                                                   #SUBSEQUENT_ENCODING:  // Statement section case 2 to 4
                                                       FOR #tempLoopCounter := #statClientIdPos TO LEN(#clientIdentifier) DO
                                                           "LMQTT_ConvertToUtf8"(character := #clientIdentifier[#tempLoopCounter],
                                                                                 convertedUtf8 => #tempConvertedUtf8,
                                                                                 bytesUsed => #tempBytesUsedUtf8,
                                                                                 error => #tempErrorConvertUtf8,
                                                                                 status => #tempStatusConvertUtf8);
                                                           IF #statSendBufferPos + #tempBytesUsedUtf8 <= #MAX_BUFFER_LEN_SEND THEN
                                                               #statClientIdPos += 1;
                                                               CASE #tempBytesUsedUtf8 OF
                                                                   #UTF_1_BYTE_USED:  // Statement section case 1
                                                                       #statSendBuffer[#statSendBufferPos] := #tempConvertedUtf8.%B0;
                                                                       #statSendBufferPos += 1;
                                                                   #UTF_2_BYTE_USED:
                                                                       #statSendBuffer[#statSendBufferPos] := #tempConvertedUtf8.%B0;
                                                                       #statSendBufferPos += 1;
                                                                       #statSendBuffer[#statSendBufferPos] := #tempConvertedUtf8.%B1;
                                                                       #statSendBufferPos += 1;
                                                                   #UTF_3_BYTE_USED:  // Statement section case 2 to 4
                                                                       #statSendBuffer[#statSendBufferPos] := #tempConvertedUtf8.%B0;
                                                                       #statSendBufferPos += 1;
                                                                       #statSendBuffer[#statSendBufferPos] := #tempConvertedUtf8.%B1;
                                                                       #statSendBufferPos += 1;
                                                                       #statSendBuffer[#statSendBufferPos] := #tempConvertedUtf8.%B2;
                                                                       #statSendBufferPos += 1;
                                                                   ELSE  // Statement section ELSE
                                                                       ;
                                                               END_CASE;
                                                           ELSE
                                                               // When buffer full
                                                               EXIT;
                                                           END_IF;
                                                       END_FOR;
                                                       IF #statClientIdPos >= LEN(#clientIdentifier) THEN
                                                           #statClientIdEncodeState := #ENCODE_DONE;
                                                       END_IF;
                                                   ELSE  // Statement section ELSE
                                                       ; // IDLE / SKIP
                                               END_CASE;
                                           END_IF;

                                           // Will Topic
                                           // If the Will Flag is set to 1, the Will Topic is the next field in the payload. It must be > 0 Bytes

                                           IF #statClientIdEncodeState = #ENCODE_DONE
                                               AND #statSendBufferPos <= #MAX_BUFFER_LEN_SEND - #TWO_BYTE_LEN_INFO THEN
                                               // When Client Id is encoded and buffer not full
                                               // And willTopic is used
                                               CASE #statWillTopicEncodeState OF
                                                   #FIRST_ENCODING:  // Statement section case 1
                                                       // ADD len info into packet

                                                       #tempWordForSliceAddress := UINT_TO_WORD(#statWillTopicLenUtf8Encoded);
                                                       #statSendBuffer[#statSendBufferPos] := #tempWordForSliceAddress.%B1; // MSB
                                                       #statSendBufferPos += 1;
                                                       #statSendBuffer[#statSendBufferPos] := #tempWordForSliceAddress.%B0; // LSB
                                                       #statSendBufferPos += 1;

                                                       FOR #tempLoopCounter := #statWillTopicPos TO LEN(#willtopic) DO
                                                           "LMQTT_ConvertToUtf8"(character := #willtopic[#tempLoopCounter],
                                                                                 convertedUtf8 => #tempConvertedUtf8,
                                                                                 bytesUsed => #tempBytesUsedUtf8,
                                                                                 error => #tempErrorConvertUtf8,
                                                                                 status => #tempStatusConvertUtf8);

                                                           IF #statSendBufferPos + #tempBytesUsedUtf8 <= #MAX_BUFFER_LEN_SEND THEN
                                                               // Increment when successful
                                                               #statWillTopicPos += 1;

                                                               CASE #tempBytesUsedUtf8 OF
                                                                   #UTF_1_BYTE_USED:  // Statement section case 1
                                                                       #statSendBuffer[#statSendBufferPos] := #tempConvertedUtf8.%B0;
                                                                       #statSendBufferPos += 1;
                                                                   #UTF_2_BYTE_USED:
                                                                       #statSendBuffer[#statSendBufferPos] := #tempConvertedUtf8.%B0;
                                                                       #statSendBufferPos += 1;
                                                                       #statSendBuffer[#statSendBufferPos] := #tempConvertedUtf8.%B1;
                                                                       #statSendBufferPos += 1;
                                                                   #UTF_3_BYTE_USED:  // Statement section case 2 to 4
                                                                       #statSendBuffer[#statSendBufferPos] := #tempConvertedUtf8.%B0;
                                                                       #statSendBufferPos += 1;
                                                                       #statSendBuffer[#statSendBufferPos] := #tempConvertedUtf8.%B1;
                                                                       #statSendBufferPos += 1;
                                                                       #statSendBuffer[#statSendBufferPos] := #tempConvertedUtf8.%B2;
                                                                       #statSendBufferPos += 1;
                                                                   ELSE  // Statement section ELSE
                                                                       ;
                                                               END_CASE;
                                                           ELSE
                                                               // When buffer full
                                                               #statWillTopicEncodeState := #SUBSEQUENT_ENCODING;
                                                               EXIT;
                                                           END_IF;
                                                       END_FOR;

                                                       IF #statWillTopicPos >= LEN(#willtopic) THEN
                                                           #statWillTopicEncodeState := #ENCODE_DONE;
                                                       END_IF;

                                                   #SUBSEQUENT_ENCODING:  // Statement section case 2 to 4
                                                       FOR #tempLoopCounter := #statWillTopicPos TO LEN(#willtopic) DO
                                                           "LMQTT_ConvertToUtf8"(character := #willtopic[#tempLoopCounter],
                                                                                 convertedUtf8 => #tempConvertedUtf8,
                                                                                 bytesUsed => #tempBytesUsedUtf8,
                                                                                 error => #tempErrorConvertUtf8,
                                                                                 status => #tempStatusConvertUtf8);

                                                           IF #statSendBufferPos + #tempBytesUsedUtf8 <= #MAX_BUFFER_LEN_SEND THEN
                                                               #statWillTopicPos += 1;
                                                               CASE #tempBytesUsedUtf8 OF
                                                                   #UTF_1_BYTE_USED:  // Statement section case 1
                                                                       #statSendBuffer[#statSendBufferPos] := #tempConvertedUtf8.%B0;
                                                                       #statSendBufferPos += 1;
                                                                   #UTF_2_BYTE_USED:
                                                                       #statSendBuffer[#statSendBufferPos] := #tempConvertedUtf8.%B0;
                                                                       #statSendBufferPos += 1;
                                                                       #statSendBuffer[#statSendBufferPos] := #tempConvertedUtf8.%B1;
                                                                       #statSendBufferPos += 1;
                                                                   #UTF_3_BYTE_USED:  // Statement section case 2 to 4
                                                                       #statSendBuffer[#statSendBufferPos] := #tempConvertedUtf8.%B0;
                                                                       #statSendBufferPos += 1;
                                                                       #statSendBuffer[#statSendBufferPos] := #tempConvertedUtf8.%B1;
                                                                       #statSendBufferPos += 1;
                                                                       #statSendBuffer[#statSendBufferPos] := #tempConvertedUtf8.%B2;
                                                                       #statSendBufferPos += 1;
                                                                   ELSE  // Statement section ELSE
                                                                       ;
                                                               END_CASE;
                                                           ELSE
                                                               // When buffer full
                                                               EXIT;
                                                           END_IF;
                                                       END_FOR;
                                                       IF #statWillTopicPos >= LEN(#willtopic) THEN
                                                           #statWillTopicEncodeState := #ENCODE_DONE;
                                                       END_IF;

                                                   ELSE  // Statement section ELSE
                                                       ;
                                               END_CASE;
                                           END_IF;

                                           // Will Message
                                           // This field consists OF a two Byte length followed BY the payload FOR the Will message expressed as a sequence bytes.

                                           IF #statClientIdEncodeState = #ENCODE_DONE
                                               AND #statWillTopicEncodeState = #ENCODE_DONE
                                               AND #statSendBufferPos <= #MAX_BUFFER_LEN_SEND - #TWO_BYTE_LEN_INFO THEN
                                               // When Client Id is encoded and buffer not full
                                               CASE #statWillMessageEncodeState OF
                                                   #FIRST_ENCODING:  // Statement section case 1
                                                       // ADD len info into packet

                                                       #tempWordForSliceAddress := UINT_TO_WORD(#statWillMessageCnt);
                                                       #statSendBuffer[#statSendBufferPos] := #tempWordForSliceAddress.%B1; // MSB
                                                       #statSendBufferPos += 1;
                                                       #statSendBuffer[#statSendBufferPos] := #tempWordForSliceAddress.%B0; // LSB
                                                       #statSendBufferPos += 1;

                                                       #tempLowerWillMsgArrayBoundary := LOWER_BOUND(ARR := #willMsgPayload, DIM := #ONE_DIMENSION);

                                                       IF #statWillMessageCnt > 0 THEN // will message exists
                                                           FOR #tempLoopCounter := #statWillMessagePos TO UINT_TO_DINT(#statWillMessageCnt - 1) DO
                                                               IF #statSendBufferPos <= #MAX_BUFFER_LEN_SEND THEN
                                                                   #statSendBuffer[#statSendBufferPos] := #willMsgPayload[#tempLowerWillMsgArrayBoundary + #tempLoopCounter];
                                                                   #statSendBufferPos += 1;
                                                                   // Increment when successful
                                                                   #statWillMessagePos += 1;
                                                               ELSE
                                                                   // When buffer full
                                                                   #statWillMessageEncodeState := #SUBSEQUENT_ENCODING;
                                                                   EXIT;
                                                               END_IF;
                                                           END_FOR;
                                                       END_IF;

                                                       // If everything was copied successfull
                                                       IF #statWillMessagePos >= #statWillMessageCnt THEN
                                                           #statWillMessageEncodeState := #ENCODE_DONE;
                                                       END_IF;

                                                   #SUBSEQUENT_ENCODING:  // Statement section case 2 to 4
                                                       #tempLowerWillMsgArrayBoundary := LOWER_BOUND(ARR := #willMsgPayload, DIM := #ONE_DIMENSION);

                                                       FOR #tempLoopCounter := #statWillMessagePos TO UINT_TO_DINT(#statWillMessageCnt - 1) DO
                                                           IF #statSendBufferPos <= #MAX_BUFFER_LEN_SEND THEN
                                                               #statSendBuffer[#statSendBufferPos] := #willMsgPayload[#tempLowerWillMsgArrayBoundary + #tempLoopCounter];
                                                               #statSendBufferPos += 1;
                                                               // Increment when successful
                                                               #statWillMessagePos += 1;
                                                           ELSE
                                                               // When Buffer Full
                                                               EXIT;
                                                           END_IF;
                                                       END_FOR;
                                                       // If everything was copied successfull
                                                       IF #statWillMessagePos >= #statWillMessageCnt THEN
                                                           #statWillMessageEncodeState := #ENCODE_DONE;
                                                       END_IF;


                                                   ELSE  // Statement section ELSE
                                                       ;
                                               END_CASE;
                                           END_IF;

                                           // Username
                                           // If the Username Flag is set to 1, the Username the next field in the payload. It must be > 0 Bytes

                                           IF #statClientIdEncodeState = #ENCODE_DONE
                                               AND (#statWillTopicEncodeState = #ENCODE_DONE OR #statWillTopicEncodeState = #NOT_USED_NO_ENCODING)
                                               AND (#statWillMessageEncodeState = #ENCODE_DONE OR #statWillTopicEncodeState = #NOT_USED_NO_ENCODING)
                                               AND #statSendBufferPos <= #MAX_BUFFER_LEN_SEND - #TWO_BYTE_LEN_INFO THEN
                                               // When Will Topic and Will Message is encoded and buffer not full
                                               CASE #statUserNameEncodeState OF
                                                   #FIRST_ENCODING:  // Statement section case 1
                                                       // ADD len info into packet

                                                       #tempWordForSliceAddress := UINT_TO_WORD(#statUsernameLenUtf8Encoded);
                                                       #statSendBuffer[#statSendBufferPos] := #tempWordForSliceAddress.%B1; // MSB
                                                       #statSendBufferPos += 1;
                                                       #statSendBuffer[#statSendBufferPos] := #tempWordForSliceAddress.%B0; // LSB
                                                       #statSendBufferPos += 1;

                                                       FOR #tempLoopCounter := #statUserNamePos TO LEN(#username) DO
                                                           "LMQTT_ConvertToUtf8"(character := #username[#tempLoopCounter],
                                                                                 convertedUtf8 => #tempConvertedUtf8,
                                                                                 bytesUsed => #tempBytesUsedUtf8,
                                                                                 error => #tempErrorConvertUtf8,
                                                                                 status => #tempStatusConvertUtf8);

                                                           IF #statSendBufferPos + #tempBytesUsedUtf8 <= #MAX_BUFFER_LEN_SEND THEN
                                                               // Increment when successful
                                                               #statUserNamePos += 1;

                                                               CASE #tempBytesUsedUtf8 OF
                                                                   #UTF_1_BYTE_USED:  // Statement section case 1
                                                                       #statSendBuffer[#statSendBufferPos] := #tempConvertedUtf8.%B0;
                                                                       #statSendBufferPos += 1;
                                                                   #UTF_2_BYTE_USED:
                                                                       #statSendBuffer[#statSendBufferPos] := #tempConvertedUtf8.%B0;
                                                                       #statSendBufferPos += 1;
                                                                       #statSendBuffer[#statSendBufferPos] := #tempConvertedUtf8.%B1;
                                                                       #statSendBufferPos += 1;
                                                                   #UTF_3_BYTE_USED:  // Statement section case 2 to 4
                                                                       #statSendBuffer[#statSendBufferPos] := #tempConvertedUtf8.%B0;
                                                                       #statSendBufferPos += 1;
                                                                       #statSendBuffer[#statSendBufferPos] := #tempConvertedUtf8.%B1;
                                                                       #statSendBufferPos += 1;
                                                                       #statSendBuffer[#statSendBufferPos] := #tempConvertedUtf8.%B2;
                                                                       #statSendBufferPos += 1;
                                                                   ELSE  // Statement section ELSE
                                                                       ;
                                                               END_CASE;
                                                           ELSE
                                                               // When buffer full
                                                               #statUserNameEncodeState := #SUBSEQUENT_ENCODING;
                                                               EXIT;
                                                           END_IF;
                                                       END_FOR;

                                                       IF #statUserNamePos >= LEN(#username) THEN
                                                           #statUserNameEncodeState := #ENCODE_DONE;
                                                       END_IF;

                                                   #SUBSEQUENT_ENCODING:  // Statement section case 2 to 4
                                                       FOR #tempLoopCounter := #statUserNamePos TO LEN(#username) DO
                                                           "LMQTT_ConvertToUtf8"(character := #username[#tempLoopCounter],
                                                                                 convertedUtf8 => #tempConvertedUtf8,
                                                                                 bytesUsed => #tempBytesUsedUtf8,
                                                                                 error => #tempErrorConvertUtf8,
                                                                                 status => #tempStatusConvertUtf8);

                                                           IF #statSendBufferPos + #tempBytesUsedUtf8 <= #MAX_BUFFER_LEN_SEND THEN
                                                               #statUserNamePos += 1;
                                                               CASE #tempBytesUsedUtf8 OF
                                                                   #UTF_1_BYTE_USED:  // Statement section case 1
                                                                       #statSendBuffer[#statSendBufferPos] := #tempConvertedUtf8.%B0;
                                                                       #statSendBufferPos += 1;
                                                                   #UTF_2_BYTE_USED:
                                                                       #statSendBuffer[#statSendBufferPos] := #tempConvertedUtf8.%B0;
                                                                       #statSendBufferPos += 1;
                                                                       #statSendBuffer[#statSendBufferPos] := #tempConvertedUtf8.%B1;
                                                                       #statSendBufferPos += 1;
                                                                   #UTF_3_BYTE_USED:  // Statement section case 2 to 4
                                                                       #statSendBuffer[#statSendBufferPos] := #tempConvertedUtf8.%B0;
                                                                       #statSendBufferPos += 1;
                                                                       #statSendBuffer[#statSendBufferPos] := #tempConvertedUtf8.%B1;
                                                                       #statSendBufferPos += 1;
                                                                       #statSendBuffer[#statSendBufferPos] := #tempConvertedUtf8.%B2;
                                                                       #statSendBufferPos += 1;
                                                                   ELSE  // Statement section ELSE
                                                                       ;
                                                               END_CASE;
                                                           ELSE
                                                               // When buffer full
                                                               EXIT;
                                                           END_IF;
                                                       END_FOR;
                                                       IF #statUserNamePos >= LEN(#username) THEN
                                                           #statUserNameEncodeState := #ENCODE_DONE;
                                                       END_IF;

                                                   ELSE  // Statement section ELSE
                                                       ;
                                               END_CASE;
                                           END_IF;

                                           // Password
                                           // If the Password Flag is set to 1, the Password the next field in the payload. It must be > 0 Bytes
                                           // Password field contains 0 to 65535 bytes OF binary data prefixed with a two Byte length field which indicates the number OF bytes used

                                           IF #statClientIdEncodeState = #ENCODE_DONE
                                               AND (#statWillTopicEncodeState = #ENCODE_DONE OR #statWillTopicEncodeState = #NOT_USED_NO_ENCODING)
                                               AND (#statWillMessageEncodeState = #ENCODE_DONE OR #statWillMessageEncodeState = #NOT_USED_NO_ENCODING)
                                               AND (#statUserNameEncodeState = #ENCODE_DONE OR #statUserNameEncodeState = #NOT_USED_NO_ENCODING)
                                               AND #statSendBufferPos <= #MAX_BUFFER_LEN_SEND - #TWO_BYTE_LEN_INFO THEN
                                               // When Will Topic and Will Message is encoded and buffer not full
                                               CASE #statPasswordEncodeState OF
                                                   #FIRST_ENCODING:  // Statement section case 1
                                                       // ADD len info into packet

                                                       #tempWordForSliceAddress := UINT_TO_WORD(#statPasswordLenUtf8Encoded);
                                                       #statSendBuffer[#statSendBufferPos] := #tempWordForSliceAddress.%B1; // MSB
                                                       #statSendBufferPos += 1;
                                                       #statSendBuffer[#statSendBufferPos] := #tempWordForSliceAddress.%B0; // LSB
                                                       #statSendBufferPos += 1;

                                                       FOR #tempLoopCounter := #statPasswordPos TO LEN(#password) DO
                                                           "LMQTT_ConvertToUtf8"(character := #password[#tempLoopCounter],
                                                                                 convertedUtf8 => #tempConvertedUtf8,
                                                                                 bytesUsed => #tempBytesUsedUtf8,
                                                                                 error => #tempErrorConvertUtf8,
                                                                                 status => #tempStatusConvertUtf8);

                                                           IF #statSendBufferPos + #tempBytesUsedUtf8 <= #MAX_BUFFER_LEN_SEND THEN
                                                               // Increment when successful
                                                               #statPasswordPos += 1;

                                                               CASE #tempBytesUsedUtf8 OF
                                                                   #UTF_1_BYTE_USED:  // Statement section case 1
                                                                       #statSendBuffer[#statSendBufferPos] := #tempConvertedUtf8.%B0;
                                                                       #statSendBufferPos += 1;
                                                                   #UTF_2_BYTE_USED:
                                                                       #statSendBuffer[#statSendBufferPos] := #tempConvertedUtf8.%B0;
                                                                       #statSendBufferPos += 1;
                                                                       #statSendBuffer[#statSendBufferPos] := #tempConvertedUtf8.%B1;
                                                                       #statSendBufferPos += 1;
                                                                   #UTF_3_BYTE_USED:  // Statement section case 2 to 4
                                                                       #statSendBuffer[#statSendBufferPos] := #tempConvertedUtf8.%B0;
                                                                       #statSendBufferPos += 1;
                                                                       #statSendBuffer[#statSendBufferPos] := #tempConvertedUtf8.%B1;
                                                                       #statSendBufferPos += 1;
                                                                       #statSendBuffer[#statSendBufferPos] := #tempConvertedUtf8.%B2;
                                                                       #statSendBufferPos += 1;
                                                                   ELSE  // Statement section ELSE
                                                                       ;
                                                               END_CASE;
                                                           ELSE
                                                               // When buffer full
                                                               #statPasswordEncodeState := #SUBSEQUENT_ENCODING;
                                                               EXIT;
                                                           END_IF;
                                                       END_FOR;

                                                       IF #statPasswordPos >= LEN(#password) THEN
                                                           #statPasswordEncodeState := #ENCODE_DONE;
                                                       END_IF;

                                                   #SUBSEQUENT_ENCODING:  // Statement section case 2 to 4
                                                       FOR #tempLoopCounter := #statPasswordPos TO LEN(#password) DO
                                                           "LMQTT_ConvertToUtf8"(character := #password[#tempLoopCounter],
                                                                                 convertedUtf8 => #tempConvertedUtf8,
                                                                                 bytesUsed => #tempBytesUsedUtf8,
                                                                                 error => #tempErrorConvertUtf8,
                                                                                 status => #tempStatusConvertUtf8);

                                                           IF #statSendBufferPos + #tempBytesUsedUtf8 <= #MAX_BUFFER_LEN_SEND THEN
                                                               #statPasswordPos += 1;
                                                               CASE #tempBytesUsedUtf8 OF
                                                                   #UTF_1_BYTE_USED:  // Statement section case 1
                                                                       #statSendBuffer[#statSendBufferPos] := #tempConvertedUtf8.%B0;
                                                                       #statSendBufferPos += 1;
                                                                   #UTF_2_BYTE_USED:
                                                                       #statSendBuffer[#statSendBufferPos] := #tempConvertedUtf8.%B0;
                                                                       #statSendBufferPos += 1;
                                                                       #statSendBuffer[#statSendBufferPos] := #tempConvertedUtf8.%B1;
                                                                       #statSendBufferPos += 1;
                                                                   #UTF_3_BYTE_USED:  // Statement section case 2 to 4
                                                                       #statSendBuffer[#statSendBufferPos] := #tempConvertedUtf8.%B0;
                                                                       #statSendBufferPos += 1;
                                                                       #statSendBuffer[#statSendBufferPos] := #tempConvertedUtf8.%B1;
                                                                       #statSendBufferPos += 1;
                                                                       #statSendBuffer[#statSendBufferPos] := #tempConvertedUtf8.%B2;
                                                                       #statSendBufferPos += 1;
                                                                   ELSE  // Statement section ELSE
                                                                       ;
                                                               END_CASE;
                                                           ELSE
                                                               // When buffer full
                                                               EXIT;
                                                           END_IF;
                                                       END_FOR;
                                                       IF #statPasswordPos >= LEN(#password) THEN
                                                           #statPasswordEncodeState := #ENCODE_DONE;
                                                       END_IF;

                                                   ELSE  // Statement section ELSE
                                                       ;
                                               END_CASE;
                                           END_IF;

                                           // set Sendlen for TSendC Block
                                           #statTsendcLen := #statSendBufferPos; // Buffer pos equals amount of elements in send array
                                           // reset buffer pos
                                           #statSendBufferPos := 0;
                                           // enable Send Req
                                           #statTsendcReq := TRUE;
                                           // Set Watchdog
                                           #statEnableTimerCommandWatchdog := TRUE;
                                           // wait for send to be done
                                           #statMqttConnectState := #MQTT_CONNECT_STATE_SEND_PACKET_WAIT_FOR_CONNACK;
                                       END_IF;
                                   END_REGION BUILD_CONNECT_PACKET

                               #MQTT_CONNECT_STATE_SEND_PACKET_WAIT_FOR_CONNACK:
                                   REGION SEND_CONNECT_PACKET_WAIT_FOR_CONNACK
                                       // check tsend status
                                       IF NOT #tempTsendcBusy AND #tempTsendcStatus = #TSENDC_JOB_DONE THEN
                                           IF (#statClientIdEncodeState = #ENCODE_DONE OR #statClientIdEncodeState = #NOT_USED_NO_ENCODING)
                                               AND (#statWillTopicEncodeState = #ENCODE_DONE OR #statWillTopicEncodeState = #NOT_USED_NO_ENCODING)
                                               AND (#statWillMessageEncodeState = #ENCODE_DONE OR #statWillMessageEncodeState = #NOT_USED_NO_ENCODING)
                                               AND (#statUserNameEncodeState = #ENCODE_DONE OR #statUserNameEncodeState = #NOT_USED_NO_ENCODING)
                                               AND (#statPasswordEncodeState = #ENCODE_DONE OR #statPasswordEncodeState = #NOT_USED_NO_ENCODING) THEN
                                               // Encoding done all sent
                                               #statPacketHeaderEncodeDone := FALSE;
                                           ELSE
                                               // More to Encode and send
                                               #statEnableTimerCommandWatchdog := FALSE;
                                               #statMqttConnectState := #MQTT_CONNECT_STATE_BUILD_PACKET;
                                           END_IF;
                                       END_IF;

                                       // Check Connect ACK packet
                                       CASE #tempMqttConnAckRcvStatus OF
                                           #NO_RESPONSE:  // IDLE
                                               // Check watchdog
                                               IF #instTimerCommandWatchdog.Q THEN
                                                   #statEnableTimerCommandWatchdog := FALSE;
                                                   #statPacketHeaderEncodeDone := FALSE;
                                                   #statStatus := #ERR_MQTT_CONNECT_TIMEOUT; // Set correct status that identifies error clearly
                                                   #statSubfunctionStatus := #ERR_MQTT_CONNECT_TIMEOUT; // Status or return value of called FBs, FCs and system blocks
                                                   #statFBErrorState := #statFBState; // Set error state number for diagnostic 
                                                   #statErrorAutoCleared := TRUE;
                                                   #statMqttConnectState := #MQTT_CONNECT_STATE_BUILD_PACKET;
                                               END_IF;
                                           #RESPONSE_GOOD:
                                               // disable watchdog
                                               #statEnableTimerCommandWatchdog := FALSE;
                                               // Encoding done all sent
                                               #statPacketHeaderEncodeDone := FALSE;
                                               // Go to Connected
                                               #statMqttConnectState := #MQTT_CONNECT_STATE_CONNECTED;
                                               #statStatus := #STATUS_MQTT_CONNECTED;
                                       END_CASE;
                                   END_REGION REGION SEND_CONNECT_PACKET

                               #MQTT_CONNECT_STATE_CONNECTED:
                                   REGION CONNECTED
                                       // Check Rising edge of input commands
                                       #tempCommandInput.%X0 := #tempPublish AND NOT #statPublishOld;
                                       #tempCommandInput.%X1 := #tempSubscribe AND NOT #statSubscribeOld;
                                       #tempCommandInput.%X2 := #tempUnsubscribe AND NOT #statUnsubscribeOld;

                                       // Start the keepalive timer if used
                                       #statEnableMqttKeepAliveTimer := #statMqttKeepAliveUsed;

                                       // set status to connected after successfully executed job
                                       IF #statStatus = #STATUS_JOB_EXECUTED THEN
                                           #statStatus := #STATUS_MQTT_CONNECTED;
                                       END_IF;

                                       // Reset done bit
                                       IF #statDone = TRUE
                                           AND #tempPublish = FALSE
                                           AND #tempSubscribe = FALSE
                                           AND #tempUnsubscribe = FALSE
                                       THEN
                                           #statDone := FALSE;
                                       END_IF;

                                       REGION MQTT_COMMANDS
                                           // When state machine is ready for a new input then assign correct command
                                           // Ping job can be overwritten by a command.
                                           IF #tempCommandInput <> #NO_COMMAND
                                               AND (#statMqttCommandState = #MQTT_COMMAND_STATE_NO_PROCESSING OR #statMqttCommandState = #MQTT_COMMAND_STATE_SEND_PING)
                                           THEN
                                               // New Input set, reset done flag
                                               #statDone := FALSE;
                                               #statMqttCommandState := BYTE_TO_DINT(#tempCommandInput);
                                           END_IF;

                                           CASE #statMqttCommandState OF
                                               #MQTT_COMMAND_STATE_NO_PROCESSING:
                                                   // EMPTY STATE
                                                   ;
                                               #MQTT_COMMAND_STATE_BUILD_PUBLISH:  // Statement section case 1
                                                   REGION PUBLISH_TO_TOPIC
                                                       // Remaining Length is the length of the variable header (TOPIC NAME + PacketID) plus the length of the Payload. 
                                                       // Max Len of Mqtt packets is per Standard 268,435,455 Bytes (ff,ff,ff,7f)
                                                       // Calculate Remain Len will be
                                                       // Len of TOPIC   (max 3*16382 WChars= 49.146 Bytes)
                                                       // plus Len of PacketID (2 Bytes)
                                                       // plus Len of Payload (max 268,435,455 - 49.146 - 2 = 268.386.307 Bytes ca. 268 MB)
                                                       // Max Array / DB Len in TIA portal is around 16 MB or 16.777.216 Byte
                                                       // Set Status
                                                       #statStatus := #STATUS_MQTT_PUBLISH;

                                                       // Must obey, if not currently sending PubAck Msg on a subscription
                                                       // Else, try in the next cycle
                                                       IF #tempTsendcBusy = FALSE // when tsendC is ready
                                                           AND #tempTsendcDone = FALSE // tsendC did not finish in this cycle
                                                           AND #statTsendcReq = FALSE // TsendC request was not already requested by pub ack msg
                                                       THEN
                                                           IF #statPacketHeaderEncodeDone = FALSE THEN

                                                               // Init
                                                               #statSendPacketTotalRemLen := 0;
                                                               #statSendBufferPos := 0;
                                                               #statPublishQos := #qos;
                                                               #statPublishMessageCnt := #publishMsgLen;
                                                               #statPublishTopicEncodeState := #FIRST_ENCODING;
                                                               #statPublishTopicPos := #FIRST_CHARACTER;
                                                               #statPublishTopicLenUtf8Encoded := 0;
                                                               #statPacketId += 1;// increment
                                                               IF (#statPacketId = 0) THEN
                                                                   #statPacketId := 1;
                                                               END_IF;
                                                               #statPacketIdEncoded := FALSE;
                                                               #statPublishEncodeMessageState := #SUBSEQUENT_ENCODING; // No len info necessary so start directly at subsequent.
                                                               #statPublishMessagePos := 0; // first array element

                                                               // verify PayloadLen
                                                               #tempMaxPublishDataArrayLen := ABS(UPPER_BOUND(ARR := #publishMsgPayload, DIM := #ONE_DIMENSION) - LOWER_BOUND(ARR := #publishMsgPayload, DIM := #ONE_DIMENSION)) + #ARRAY_LEN_OFFSET_PLUS_1;

                                                               // check necessary boundaries
                                                               IF #tempMaxPublishDataArrayLen < #statPublishMessageCnt THEN
                                                                   #statStatus := #ERR_CNT_EXCEEDS_ARRAY_DIMENSION; // Set correct status that identifies error clearly
                                                                   #statSubfunctionStatus := #ERR_CNT_EXCEEDS_ARRAY_DIMENSION; // Status or return value of called FBs, FCs and system blocks
                                                                   #statFBErrorState := #statFBState; // Set error state number for diagnostic 
                                                                   #statErrorAutoCleared := TRUE;
                                                                   #statMqttCommandState := #MQTT_COMMAND_STATE_NO_PROCESSING;
                                                               ELSIF LEN(#mqttTopic) = #LEN_NULL THEN
                                                                   #statStatus := #ERR_MQTT_COMMAND_PUBLISH_TOPIC_INVALID; // Set correct status that identifies error clearly
                                                                   #statSubfunctionStatus := #ERR_MQTT_COMMAND_PUBLISH_TOPIC_INVALID; // Status or return value of called FBs, FCs and system blocks
                                                                   #statFBErrorState := #statFBState; // Set error state number for diagnostic 
                                                                   #statErrorAutoCleared := TRUE;
                                                                   #statMqttCommandState := #MQTT_COMMAND_STATE_NO_PROCESSING;
                                                               ELSIF #statPublishQos > #MQTT_QOS_2 THEN
                                                                   #statStatus := #ERR_QOS_INVALID; // Set correct status that identifies error clearly
                                                                   #statSubfunctionStatus := #ERR_QOS_INVALID; // Status or return value of called FBs, FCs and system blocks
                                                                   #statFBErrorState := #statFBState; // Set error state number for diagnostic 
                                                                   #statErrorAutoCleared := TRUE;
                                                                   #statMqttCommandState := #MQTT_COMMAND_STATE_NO_PROCESSING;
                                                               ELSE // All ok
                                                                   // Add amount of bytes for publish message
                                                                   #statSendPacketTotalRemLen := #statSendPacketTotalRemLen + #statPublishMessageCnt;
                                                                   // add publish  topic len
                                                                   FOR #tempLoopCounter := #FIRST_CHARACTER TO LEN(#mqttTopic) DO
                                                                       "LMQTT_ConvertToUtf8"(character := #mqttTopic[#tempLoopCounter],
                                                                                             convertedUtf8 => #tempConvertedUtf8,
                                                                                             bytesUsed => #tempBytesUsedUtf8,
                                                                                             error => #tempErrorConvertUtf8,
                                                                                             status => #tempStatusConvertUtf8);
                                                                       #statPublishTopicLenUtf8Encoded := #statPublishTopicLenUtf8Encoded + #tempBytesUsedUtf8;
                                                                   END_FOR;
                                                                   #statSendPacketTotalRemLen := #statSendPacketTotalRemLen + #statPublishTopicLenUtf8Encoded + #TWO_BYTE_LEN_INFO;

                                                                   // Build Publish Telegram
                                                                   // Fixed Header - Write Packet Type
                                                                   #statSendBuffer[#statSendBufferPos] := #MQTT_MSG_TYPE_PUBLISH;
                                                                   // Set DUP flag always to FALSE
                                                                   #statSendBuffer[#statSendBufferPos].%X3 := FALSE;
                                                                   // Set QoS Level
                                                                   CASE #statPublishQos OF
                                                                       #MQTT_QOS_0:  // Statement section case 0
                                                                           #statSendBuffer[#statSendBufferPos] := #statSendBuffer[#statSendBufferPos] OR #MQTT_MSG_QOS0;
                                                                       #MQTT_QOS_1:  // Statement section case 1
                                                                           #statSendBuffer[#statSendBufferPos] := #statSendBuffer[#statSendBufferPos] OR #MQTT_MSG_QOS1;
                                                                           // Add two byte len info for Mandatory packet ID
                                                                           #statSendPacketTotalRemLen := #statSendPacketTotalRemLen + #TWO_BYTE_LEN_INFO;
                                                                       #MQTT_QOS_2: // Statement section case 2
                                                                           #statSendBuffer[#statSendBufferPos] := #statSendBuffer[#statSendBufferPos] OR #MQTT_MSG_QOS2;
                                                                           // Add two byte len info for Mandatory packet ID
                                                                           #statSendPacketTotalRemLen := #statSendPacketTotalRemLen + #TWO_BYTE_LEN_INFO;
                                                                       ELSE
                                                                           ;
                                                                   END_CASE;
                                                                   // Set retain bit
                                                                   #statSendBuffer[#statSendBufferPos].%X0 := #retain;

                                                                   #statSendBufferPos += 1; // increment

                                                                   // Write Remaining Packet Len info 
                                                                   WHILE (#statSendPacketTotalRemLen > #DEFAULT_VALUE_ZERO)
                                                                   DO// See MQTT Spec for explanation of this calculation
                                                                       #statEncodedRemPacketLenAsByte := UDINT_TO_BYTE(#statSendPacketTotalRemLen MOD #SEND_LEN_MULTIPLIER_UDINT_128);
                                                                       #statSendPacketTotalRemLen := #statSendPacketTotalRemLen / #SEND_LEN_MULTIPLIER_UDINT_128;
                                                                       // if there are more data to encode, set the top bit of this byte
                                                                       IF #statSendPacketTotalRemLen > #DEFAULT_VALUE_ZERO THEN
                                                                           // Do this and continue while loop
                                                                           #statEncodedRemPacketLenAsByte := #statEncodedRemPacketLenAsByte OR UDINT_TO_BYTE(#SEND_LEN_MULTIPLIER_UDINT_128);
                                                                           #statSendBuffer[#statSendBufferPos] := #statEncodedRemPacketLenAsByte;
                                                                           #statSendBufferPos += 1;
                                                                       ELSE
                                                                           // do this and leave while loop
                                                                           #statSendBuffer[#statSendBufferPos] := #statEncodedRemPacketLenAsByte;
                                                                           #statSendBufferPos += 1;
                                                                       END_IF;
                                                                   END_WHILE;
                                                                   // When all done, set encode to true
                                                                   #statPacketHeaderEncodeDone := TRUE;
                                                               END_IF;
                                                           END_IF;

                                                           // Header Encoded - now Topic, PacketId and Message need to be encoded.
                                                           IF #statPacketHeaderEncodeDone = TRUE THEN

                                                               // Publish Topic
                                                               IF #statSendBufferPos <= #MAX_BUFFER_LEN_SEND - #TWO_BYTE_LEN_INFO THEN
                                                                   CASE #statPublishTopicEncodeState OF
                                                                       #FIRST_ENCODING:  // Statement section case 1
                                                                           // ADD len info into packet

                                                                           #tempWordForSliceAddress := UINT_TO_WORD(#statPublishTopicLenUtf8Encoded);
                                                                           #statSendBuffer[#statSendBufferPos] := #tempWordForSliceAddress.%B1; // MSB
                                                                           #statSendBufferPos += 1;
                                                                           #statSendBuffer[#statSendBufferPos] := #tempWordForSliceAddress.%B0; // LSB
                                                                           #statSendBufferPos += 1;

                                                                           FOR #tempLoopCounter := #statPublishTopicPos TO LEN(#mqttTopic) DO
                                                                               "LMQTT_ConvertToUtf8"(character := #mqttTopic[#tempLoopCounter],
                                                                                                     convertedUtf8 => #tempConvertedUtf8,
                                                                                                     bytesUsed => #tempBytesUsedUtf8,
                                                                                                     error => #tempErrorConvertUtf8,
                                                                                                     status => #tempStatusConvertUtf8);

                                                                               IF #statSendBufferPos + #tempBytesUsedUtf8 <= #MAX_BUFFER_LEN_SEND THEN
                                                                                   #statPublishTopicPos += 1;
                                                                                   CASE #tempBytesUsedUtf8 OF
                                                                                       #UTF_1_BYTE_USED:  // Statement section case 1
                                                                                           #statSendBuffer[#statSendBufferPos] := #tempConvertedUtf8.%B0;
                                                                                           #statSendBufferPos += 1;
                                                                                       #UTF_2_BYTE_USED:
                                                                                           #statSendBuffer[#statSendBufferPos] := #tempConvertedUtf8.%B0;
                                                                                           #statSendBufferPos += 1;
                                                                                           #statSendBuffer[#statSendBufferPos] := #tempConvertedUtf8.%B1;
                                                                                           #statSendBufferPos += 1;
                                                                                       #UTF_3_BYTE_USED:  // Statement section case 2 to 4
                                                                                           #statSendBuffer[#statSendBufferPos] := #tempConvertedUtf8.%B0;
                                                                                           #statSendBufferPos += 1;
                                                                                           #statSendBuffer[#statSendBufferPos] := #tempConvertedUtf8.%B1;
                                                                                           #statSendBufferPos += 1;
                                                                                           #statSendBuffer[#statSendBufferPos] := #tempConvertedUtf8.%B2;
                                                                                           #statSendBufferPos += 1;
                                                                                       ELSE  // Statement section ELSE
                                                                                           ;
                                                                                   END_CASE;
                                                                               ELSE
                                                                                   // When buffer full
                                                                                   #statPublishTopicEncodeState := #SUBSEQUENT_ENCODING;
                                                                                   EXIT;
                                                                               END_IF;
                                                                           END_FOR;
                                                                           IF #statPublishTopicPos >= LEN(#mqttTopic) THEN
                                                                               #statPublishTopicEncodeState := #ENCODE_DONE;
                                                                           END_IF;


                                                                       #SUBSEQUENT_ENCODING:  // Statement section case 2 to 4
                                                                           FOR #tempLoopCounter := #statPublishTopicPos TO LEN(#mqttTopic) DO

                                                                               "LMQTT_ConvertToUtf8"(character := #mqttTopic[#tempLoopCounter],
                                                                                                     convertedUtf8 => #tempConvertedUtf8,
                                                                                                     bytesUsed => #tempBytesUsedUtf8,
                                                                                                     error => #tempErrorConvertUtf8,
                                                                                                     status => #tempStatusConvertUtf8);
                                                                               IF #statSendBufferPos + #tempBytesUsedUtf8 <= #MAX_BUFFER_LEN_SEND THEN
                                                                                   #statPublishTopicPos += 1;
                                                                                   CASE #tempBytesUsedUtf8 OF
                                                                                       #UTF_1_BYTE_USED:  // Statement section case 1
                                                                                           #statSendBuffer[#statSendBufferPos] := #tempConvertedUtf8.%B0;
                                                                                           #statSendBufferPos += 1;
                                                                                       #UTF_2_BYTE_USED:
                                                                                           #statSendBuffer[#statSendBufferPos] := #tempConvertedUtf8.%B0;
                                                                                           #statSendBufferPos += 1;
                                                                                           #statSendBuffer[#statSendBufferPos] := #tempConvertedUtf8.%B1;
                                                                                           #statSendBufferPos += 1;
                                                                                       #UTF_3_BYTE_USED:  // Statement section case 2 to 4
                                                                                           #statSendBuffer[#statSendBufferPos] := #tempConvertedUtf8.%B0;
                                                                                           #statSendBufferPos += 1;
                                                                                           #statSendBuffer[#statSendBufferPos] := #tempConvertedUtf8.%B1;
                                                                                           #statSendBufferPos += 1;
                                                                                           #statSendBuffer[#statSendBufferPos] := #tempConvertedUtf8.%B2;
                                                                                           #statSendBufferPos += 1;
                                                                                       ELSE  // Statement section ELSE
                                                                                           ;
                                                                                   END_CASE;
                                                                               ELSE
                                                                                   // When buffer full
                                                                                   EXIT;
                                                                               END_IF;
                                                                           END_FOR;
                                                                           IF #statPublishTopicPos >= LEN(#mqttTopic) THEN
                                                                               #statPublishTopicEncodeState := #ENCODE_DONE;
                                                                           END_IF;
                                                                       ELSE  // SKIP if done
                                                                           ;
                                                                   END_CASE;
                                                               END_IF;

                                                               // Encode MessageID, when QOS > 0 and  Topic done and buffer not full
                                                               IF #statPublishTopicEncodeState = #ENCODE_DONE
                                                                   AND #statPacketIdEncoded = FALSE
                                                                   AND #statSendBufferPos <= #MAX_BUFFER_LEN_SEND - #TWO_BYTE_LEN_INFO THEN
                                                                   // Check QoS - only necessary if QoS >0
                                                                   CASE #statPublishQos OF
                                                                       #MQTT_QOS_1:
                                                                           #tempWordForSliceAddress := UINT_TO_WORD(#statPacketId);
                                                                           #statSendBuffer[#statSendBufferPos] := #tempWordForSliceAddress.%B1; // MSB
                                                                           #statSendBufferPos += 1;
                                                                           #statSendBuffer[#statSendBufferPos] := #tempWordForSliceAddress.%B0; // LSB
                                                                           #statSendBufferPos += 1;
                                                                       #MQTT_QOS_2:
                                                                           #tempWordForSliceAddress := UINT_TO_WORD(#statPacketId);
                                                                           #statSendBuffer[#statSendBufferPos] := #tempWordForSliceAddress.%B1; // MSB
                                                                           #statSendBufferPos += 1;
                                                                           #statSendBuffer[#statSendBufferPos] := #tempWordForSliceAddress.%B0; // LSB
                                                                           #statSendBufferPos += 1;
                                                                       ELSE
                                                                           // No packet id to encode here
                                                                           ;
                                                                   END_CASE;
                                                                   // Finally:
                                                                   #statPacketIdEncoded := TRUE;
                                                               END_IF;

                                                               // Encode Payload, when  Topic done and PacketID Done and buffer not full
                                                               IF #statPublishTopicEncodeState = #ENCODE_DONE
                                                                   AND #statPacketIdEncoded = TRUE
                                                                   AND #statSendBufferPos < #MAX_BUFFER_LEN_SEND THEN

                                                                   // Publish Message Encoding
                                                                   // This Contains the payload from the publish message expressed as a sequence bytes.
                                                                   CASE #statPublishEncodeMessageState OF
                                                                       #SUBSEQUENT_ENCODING:  // Statement section case 2 to 4
                                                                           #tempLowerBoundPublishDataArray := LOWER_BOUND(ARR := #publishMsgPayload, DIM := #ONE_DIMENSION);

                                                                           FOR #tempLoopCounter := #statPublishMessagePos TO UDINT_TO_DINT(#statPublishMessageCnt - 1) DO
                                                                               IF #statSendBufferPos <= #MAX_BUFFER_LEN_SEND THEN
                                                                                   #statSendBuffer[#statSendBufferPos] := #publishMsgPayload[#tempLowerBoundPublishDataArray + #tempLoopCounter];
                                                                                   #statSendBufferPos += 1;
                                                                                   // Increment when successful
                                                                                   #statPublishMessagePos += 1;
                                                                               ELSE
                                                                                   // When Buffer Full
                                                                                   EXIT;
                                                                               END_IF;
                                                                           END_FOR;
                                                                           // If everything was copied successfull
                                                                           IF #statPublishMessagePos >= #statPublishMessageCnt THEN
                                                                               #statPublishEncodeMessageState := #ENCODE_DONE;
                                                                           END_IF;
                                                                       ELSE  // Statement section ELSE
                                                                           ;
                                                                   END_CASE;
                                                               END_IF;

                                                               // set Sendlen for TSendC Block
                                                               #statTsendcLen := #statSendBufferPos; // Buffer pos equals amount of elements in send array
                                                               // reset buffer pos
                                                               #statSendBufferPos := 0;
                                                               // enable Send Req
                                                               #statTsendcReq := TRUE;
                                                               // Set Watchdog
                                                               #statEnableTimerCommandWatchdog := TRUE;
                                                               // wait for send to be done
                                                               #statMqttCommandState := #MQTT_COMMAND_STATE_SEND_PUBLISH;
                                                           END_IF;
                                                       END_IF;
                                                   END_REGION PUBLISH_TO_TOPIC

                                               #MQTT_COMMAND_STATE_SEND_PUBLISH:
                                                   REGION SEND_PUBLISH_WAIT_FOR_RESPONSE
                                                       // check tsend status
                                                       IF NOT #tempTsendcBusy AND #tempTsendcStatus = #TSENDC_JOB_DONE THEN

                                                           IF #statPublishTopicEncodeState = #ENCODE_DONE
                                                               AND #statPublishEncodeMessageState = #ENCODE_DONE
                                                           THEN
                                                               // Encoding done all sent
                                                               #statPacketHeaderEncodeDone := FALSE;
                                                               // with QoS = 0 Job done
                                                               IF #statPublishQos = #MQTT_QOS_0 THEN
                                                                   // job done
                                                                   #statDone := TRUE;
                                                                   // go back to idle
                                                                   #statMqttCommandState := #MQTT_COMMAND_STATE_NO_PROCESSING;
                                                                   // reset Watchdog
                                                                   #statEnableTimerCommandWatchdog := FALSE;
                                                                   // Set Status back to connected
                                                                   #statStatus := #STATUS_JOB_EXECUTED;
                                                               END_IF;
                                                           ELSE
                                                               // More to Encode and send
                                                               #statEnableTimerCommandWatchdog := FALSE;
                                                               #statMqttCommandState := #MQTT_COMMAND_STATE_BUILD_PUBLISH;
                                                           END_IF;
                                                       END_IF;

                                                       // check watchdog if QoS is 1/2 and no responses have been received in this cycle
                                                       IF #instTimerCommandWatchdog.Q
                                                           AND #statPublishQos <> #MQTT_QOS_0
                                                           AND #tempMqttPubAckRcv = #NO_RESPONSE
                                                           AND #statMqttPubRecRcv = #NO_RESPONSE
                                                           AND #tempMqttPubCompRcv = #NO_RESPONSE
                                                       THEN
                                                           #statEnableTimerCommandWatchdog := FALSE;
                                                           #statStatus := #ERR_MQTT_COMMAND_SEND_TIMEOUT; // Set correct status that identifies error clearly
                                                           #statSubfunctionStatus := #ERR_MQTT_COMMAND_SEND_TIMEOUT; // Status or return value of called FBs, FCs and system blocks
                                                           #statFBErrorState := #statFBState; // Set error state number for diagnostic 
                                                           #statErrorAutoCleared := TRUE;
                                                           #statMqttCommandState := #MQTT_COMMAND_STATE_NO_PROCESSING;
                                                       END_IF;

                                                       // When QoS = 1; Wait for Publish ACK packet
                                                       CASE #tempMqttPubAckRcv OF
                                                           #NO_RESPONSE:
                                                               ;
                                                           #RESPONSE_GOOD:
                                                               // disable watchdog
                                                               #statEnableTimerCommandWatchdog := FALSE;
                                                               // Encoding done all sent
                                                               #statPacketHeaderEncodeDone := FALSE;
                                                               // Publish QoS 1 = Done
                                                               #statDone := TRUE;
                                                               #statMqttCommandState := #MQTT_COMMAND_STATE_NO_PROCESSING;
                                                               // Set Status back to connected
                                                               #statStatus := #STATUS_JOB_EXECUTED;
                                                           #RESPONSE_PACKET_ID_INVALID:
                                                               #statStatus := #ERR_MQTT_PACKET_ID_INVALID; // Set correct status that identifies error clearly
                                                               #statSubfunctionStatus := #ERR_MQTT_PACKET_ID_INVALID; // Status or return value of called FBs, FCs and system blocks
                                                               #statFBErrorState := #statFBState; // Set error state number for diagnostic 
                                                               #statErrorAutoCleared := TRUE;
                                                               #statMqttCommandState := #MQTT_COMMAND_STATE_NO_PROCESSING;
                                                       END_CASE;

                                                       // When QOS = 2 and Pub Rec Receieved:
                                                       CASE #statMqttPubRecRcv OF
                                                           #NO_RESPONSE:  // 0 IDLE
                                                               ;
                                                           #RESPONSE_GOOD:
                                                               IF #instTsendC.STATUS = #TSENDC_JOB_DONE OR #instTsendC.STATUS = #TSENDC_EST_OK THEN
                                                                   // Encoding done all sent
                                                                   #statPacketHeaderEncodeDone := FALSE;
                                                                   // Send Publish Release packet
                                                                   #statSendBufferPos := 0;
                                                                   #statSendBuffer[#statSendBufferPos] := #MQTT_MSG_TYPE_PUBREL OR #MQTT_MSG_QOS1;
                                                                   #statSendBufferPos += 1;
                                                                   // Remaining Lenght (must be 2)
                                                                   #statSendBuffer[#statSendBufferPos] := #REMAINING_LEN_2;
                                                                   #statSendBufferPos += 1;
                                                                   // add packet id 
                                                                   #tempWordForSliceAddress := UINT_TO_WORD(#statPacketId);
                                                                   #statSendBuffer[#statSendBufferPos] := #tempWordForSliceAddress.%B1; // MSB
                                                                   #statSendBufferPos += 1;
                                                                   #statSendBuffer[#statSendBufferPos] := #tempWordForSliceAddress.%B0; // LSB
                                                                   #statSendBufferPos += 1;
                                                                   #statTsendcLen := #statSendBufferPos;
                                                                   // Start send request
                                                                   #statTsendcReq := TRUE;
                                                                   #statMqttPubRecRcv := #NO_RESPONSE;

                                                                   // Reset watchdog and start
                                                                   RESET_TIMER(#instTimerCommandWatchdog);
                                                                   #statEnableTimerCommandWatchdog := TRUE;
                                                               END_IF;
                                                               // Stay in State
                                                           #RESPONSE_PACKET_ID_INVALID:
                                                               #statStatus := #ERR_MQTT_PACKET_ID_INVALID; // Set correct status that identifies error clearly
                                                               #statSubfunctionStatus := #ERR_MQTT_PACKET_ID_INVALID; // Status or return value of called FBs, FCs and system blocks
                                                               #statFBErrorState := #statFBState; // Set error state number for diagnostic 
                                                               #statErrorAutoCleared := TRUE;
                                                               #statMqttCommandState := #MQTT_COMMAND_STATE_NO_PROCESSING;
                                                       END_CASE;

                                                       // When QOS = 2 and Pub Complete Receieved:
                                                       CASE #tempMqttPubCompRcv OF
                                                           #NO_RESPONSE:  // Idle
                                                               ;
                                                           #RESPONSE_GOOD:  // When QOS = 2 and Pub Complete Receieved:
                                                               // disable watchdog
                                                               #statEnableTimerCommandWatchdog := FALSE;
                                                               // Encoding done all sent
                                                               #statPacketHeaderEncodeDone := FALSE;
                                                               // Publish QoS 2 = Done
                                                               #statDone := TRUE;

                                                               #statMqttCommandState := #MQTT_COMMAND_STATE_NO_PROCESSING;
                                                               // Set Status back to connected
                                                               #statStatus := #STATUS_JOB_EXECUTED;
                                                           #RESPONSE_PACKET_ID_INVALID:
                                                               #statStatus := #ERR_MQTT_PACKET_ID_INVALID; // Set correct status that identifies error clearly
                                                               #statSubfunctionStatus := #ERR_MQTT_PACKET_ID_INVALID; // Status or return value of called FBs, FCs and system blocks
                                                               #statFBErrorState := #statFBState; // Set error state number for diagnostic 
                                                               #statErrorAutoCleared := TRUE;
                                                               #statMqttCommandState := #MQTT_COMMAND_STATE_NO_PROCESSING;
                                                       END_CASE;
                                                   END_REGION MQTT_COMMAND_SEND_PUBLISH

                                               #MQTT_COMMAND_STATE_BUILD_SUBSCRIBE:  // Statement section case 2 
                                                   REGION SUBSCRIBE_TO_TOPIC
                                                       // Remaining Length is the length of the variable header (PacketID, 2Bytes) plus the length of the Payload. 
                                                       // Max Len of Mqtt packets is per Standard 268,435,455 Bytes (ff,ff,ff,7f)
                                                       // Calculate Remain Len will be
                                                       // Len of TOPIC   (max 3*16382 WChars= 49.146 Bytes)
                                                       // LenInfo Topic (2Byte)
                                                       // QoS of Topic (1Byte)

                                                       // Set Status
                                                       #statStatus := #STATUS_MQTT_SUBSCRIBE;
                                                       // Must obey, if not currently sending PubAck Msg on a subscription
                                                       // Else, try in the next cycle
                                                       IF #tempTsendcBusy = FALSE // when tsendC is ready
                                                           AND #tempTsendcDone = FALSE // tsendC did not finish in this cycle
                                                           AND #statTsendcReq = FALSE // TsendC request was not already requested by pub ack msg
                                                       THEN
                                                           IF #statPacketHeaderEncodeDone = FALSE THEN

                                                               // Init
                                                               #statSendPacketTotalRemLen := 0;
                                                               #statSendBufferPos := 0;
                                                               #statSubscribeQos := #qos;
                                                               #statSubscribeTopicEncodeState := #FIRST_ENCODING;
                                                               #statSubscribeTopicPos := #FIRST_CHARACTER;
                                                               #statSubscribeTopicLenUtf8Encoded := 0;
                                                               #statPacketId += 1;// increment
                                                               IF #statPacketId = 0 THEN
                                                                   #statPacketId := 1;
                                                               END_IF;
                                                               #statSubscribeQosEncoded := FALSE;

                                                               // check necessary boundaries

                                                               IF LEN(#mqttTopic) = #LEN_NULL THEN
                                                                   #statStatus := #ERR_MQTT_COMMAND_SUBSCRIBE_TOPIC_INVALID; // Set correct status that identifies error clearly
                                                                   #statSubfunctionStatus := #ERR_MQTT_COMMAND_SUBSCRIBE_TOPIC_INVALID; // Status or return value of called FBs, FCs and system blocks
                                                                   #statFBErrorState := #statFBState; // Set error state number for diagnostic 
                                                                   #statErrorAutoCleared := TRUE;
                                                                   #statMqttCommandState := #MQTT_COMMAND_STATE_NO_PROCESSING;
                                                               ELSIF #statSubscribeQos > #MQTT_QOS_2 THEN // NEW: Allow Subscribe with QoS2
                                                                   #statStatus := #ERR_QOS_INVALID; // Set correct status that identifies error clearly
                                                                   #statSubfunctionStatus := #ERR_QOS_INVALID; // Status or return value of called FBs, FCs and system blocks
                                                                   #statFBErrorState := #statFBState; // Set error state number for diagnostic 
                                                                   #statErrorAutoCleared := TRUE;
                                                                   #statMqttCommandState := #MQTT_COMMAND_STATE_NO_PROCESSING;
                                                               ELSE // All ok
                                                                   // Add two Byte for Packet ID:
                                                                   #statSendPacketTotalRemLen := #statSendPacketTotalRemLen + #TWO_BYTE_LEN_INFO;
                                                                   // Add one Byte for QoS Info:
                                                                   #statSendPacketTotalRemLen := #statSendPacketTotalRemLen + #ONE_BYTE_LEN_INFO;
                                                                   // add subscribe  topic len
                                                                   FOR #tempLoopCounter := #FIRST_CHARACTER TO LEN(#mqttTopic) DO
                                                                       "LMQTT_ConvertToUtf8"(character := #mqttTopic[#tempLoopCounter],
                                                                                             convertedUtf8 => #tempConvertedUtf8,
                                                                                             bytesUsed => #tempBytesUsedUtf8,
                                                                                             error => #tempErrorConvertUtf8,
                                                                                             status => #tempStatusConvertUtf8);
                                                                       #statSubscribeTopicLenUtf8Encoded := #statSubscribeTopicLenUtf8Encoded + #tempBytesUsedUtf8;
                                                                   END_FOR;
                                                                   // Add len of topic plus len info
                                                                   #statSendPacketTotalRemLen := #statSendPacketTotalRemLen + #statSubscribeTopicLenUtf8Encoded + #TWO_BYTE_LEN_INFO;

                                                                   // Build Subscribe Telegram
                                                                   // Fixed Header - Write Packet Type
                                                                   #statSendBuffer[#statSendBufferPos] := #MQTT_MSG_TYPE_SUBSCRIBE OR #MQTT_MSG_QOS1;
                                                                   #statSendBufferPos += 1; // increment

                                                                   // Write Remaining Packet Len info 
                                                                   WHILE (#statSendPacketTotalRemLen > #DEFAULT_VALUE_ZERO)
                                                                   DO// See MQTT Spec for explanation of this calculation
                                                                       #statEncodedRemPacketLenAsByte := UDINT_TO_BYTE(#statSendPacketTotalRemLen MOD #SEND_LEN_MULTIPLIER_UDINT_128);
                                                                       #statSendPacketTotalRemLen := #statSendPacketTotalRemLen / #SEND_LEN_MULTIPLIER_UDINT_128;
                                                                       // if there are more data to encode, set the top bit of this byte
                                                                       IF #statSendPacketTotalRemLen > #DEFAULT_VALUE_ZERO THEN
                                                                           // Do this and continue while loop
                                                                           #statEncodedRemPacketLenAsByte := #statEncodedRemPacketLenAsByte OR UDINT_TO_BYTE(#SEND_LEN_MULTIPLIER_UDINT_128);
                                                                           #statSendBuffer[#statSendBufferPos] := #statEncodedRemPacketLenAsByte;
                                                                           #statSendBufferPos += 1;
                                                                       ELSE
                                                                           // do this and leave while loop
                                                                           #statSendBuffer[#statSendBufferPos] := #statEncodedRemPacketLenAsByte;
                                                                           #statSendBufferPos += 1;
                                                                       END_IF;
                                                                   END_WHILE;

                                                                   // Set Packet Id
                                                                   #tempWordForSliceAddress := UINT_TO_WORD(#statPacketId);
                                                                   #statSendBuffer[#statSendBufferPos] := #tempWordForSliceAddress.%B1; // MSB
                                                                   #statSendBufferPos += 1;
                                                                   #statSendBuffer[#statSendBufferPos] := #tempWordForSliceAddress.%B0; // LSB
                                                                   #statSendBufferPos += 1;

                                                                   // When all done, set encode to true
                                                                   #statPacketHeaderEncodeDone := TRUE;
                                                               END_IF;
                                                           END_IF;
                                                           // Header Encoded 
                                                           IF #statPacketHeaderEncodeDone = TRUE THEN
                                                               // Header Encoded - now Topic and qos encoding
                                                               // Subscribe Topic
                                                               IF #statSendBufferPos <= #MAX_BUFFER_LEN_SEND - #TWO_BYTE_LEN_INFO THEN
                                                                   CASE #statSubscribeTopicEncodeState OF
                                                                       #FIRST_ENCODING:  // Statement section case 1
                                                                           // ADD len info into packet
                                                                           #tempWordForSliceAddress := UINT_TO_WORD(#statSubscribeTopicLenUtf8Encoded);
                                                                           #statSendBuffer[#statSendBufferPos] := #tempWordForSliceAddress.%B1; // MSB
                                                                           #statSendBufferPos += 1;
                                                                           #statSendBuffer[#statSendBufferPos] := #tempWordForSliceAddress.%B0; // LSB
                                                                           #statSendBufferPos += 1;

                                                                           FOR #tempLoopCounter := #statSubscribeTopicPos TO LEN(#mqttTopic) DO
                                                                               "LMQTT_ConvertToUtf8"(character := #mqttTopic[#tempLoopCounter],
                                                                                                     convertedUtf8 => #tempConvertedUtf8,
                                                                                                     bytesUsed => #tempBytesUsedUtf8,
                                                                                                     error => #tempErrorConvertUtf8,
                                                                                                     status => #tempStatusConvertUtf8);

